// TIA Portal V21 export
// export: Created 2026-11-10T07:35:17.7479988Z, ExportSetting WithDefaults, DisplayName Totally Integrated Automation Portal, DisplayVersion V21 Update 3, DisplayName STEP 7 Professional, DisplayVersion V21 Update 3, DisplayName STEP 7 Safety, DisplayVersion V21, DisplayName Tech WebApplication, DisplayVersion V21, DisplayName WinCC Basic/Comfort/Advanced, DisplayVersion V21 Update 3, DisplayName WinCC Unified, DisplayVersion V21 Update 3
FUNCTION_BLOCK "FB_Lad_ex130"   // FB49, LAD
{ S7_Optimized_Access := 'TRUE' }
VERSION : 0.1
// stored: AutoNumber true, IsIECCheckEnabled false, IsRetainMemResEnabled false, MemoryReserve 100, SetENOAutomatically false, UDAEnableTagReadback false
   VAR_INPUT
      v_laddr : HW_IOSYSTEM;
      v_mode : UInt;
      v_ret_val : Int;
   END_VAR
   VAR_IN_OUT
      v_state : Variant;
   END_VAR
BEGIN

REGION Network 1: DeviceStates - Read module status information in an IO system
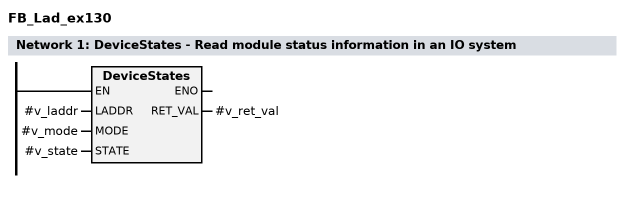
   RUNG wire#powerrail
      DeviceStates(LADDR := #v_laddr, MODE := #v_mode, Ret_Val => #v_ret_val, STATE := #v_state)
   END_RUNG
   // the same network as SCL:
   #v_ret_val := DeviceStates(LADDR := #v_laddr, MODE := #v_mode, STATE := #v_state);
END_REGION
END_FUNCTION_BLOCK
